(* IEC 61131-3 sources: plc-sbom-builder/samples/maschine-xy/programm/Roboterzelle, 1 file *)

(* ---- GVL.st ---- *)
// Globale Variablen der Roboterzelle
VAR_GLOBAL
    bNotHalt : BOOL;
END_VAR
